(*
SPDX-FileCopyrightText: c 2026 Oleksandr Tiutyk <trofimich@gmail.com>
SPDX-License-Identifier: MIT
License: https://opensource.org/license/mit
*)

(*!
<summary>Groups fixed-capacity dictionary lookup, update, removal, clear and overflow cases.</summary>
<description>
Owns the child cases, their fixed registration array and the dictionaries borrowed by the common cases.
Each borrowed fixture is reserved for its case throughout the group lifetime. Use from one task at a stable address.
</description>
*)

{attribute 'no_assign'}
{attribute 'no_explicit_call' := 'do not call this function block directly'}
FUNCTION_BLOCK StaticDictionaryTestGroup EXTENDS TOF_Testing.TestGroup<5>
VAR_STAT
	{attribute 'hide'}
	_ClassName : STRING := __POUNAME();
END_VAR
VAR
	_SetAndGetDictionary : TOF_Collections.Dictionary<7>(keyValidator := 0, valueValidator := 0, keyEqualityComparer := 0);
	_RemoveDictionary : TOF_Collections.Dictionary<7>(keyValidator := 0, valueValidator := 0, keyEqualityComparer := 0);
	_ContainsDictionary : TOF_Collections.Dictionary<7>(keyValidator := 0, valueValidator := 0, keyEqualityComparer := 0);

	_SetAndGet : DictionarySetAndGetTest(name := "SetAndGet", parent := THIS^, dictionary := _SetAndGetDictionary);
	_Remove : DictionaryRemoveTest(name := "Remove", parent := THIS^, dictionary := _RemoveDictionary);
	_Contains : DictionaryContainsTest(name := "Contains", parent := THIS^, dictionary := _ContainsDictionary);
	_Clear : StaticDictionaryClearTest(name := "Clear", parent := THIS^);
	_Overflow : StaticDictionaryOverflowTest(name := "Overflow", parent := THIS^);

	_Children : ARRAY [0.._ChildCount - 1] OF TOF_Testing.ITestElement :=
	[
		_SetAndGet,
		_Remove,
		_Contains,
		_Clear,
		_Overflow
	];
END_VAR

//! <summary>Borrows the fixed child array. Callers must not modify it.</summary>
{attribute 'monitoring' := 'call'}
PROPERTY Children : REFERENCE TO ARRAY [0.._ChildCount - 1] OF TOF_Testing.ITestElement
GET
Children REF= _Children;
END_GET
END_PROPERTY

//! <summary>Borrows the concrete class name. Callers must not modify it.</summary>
{attribute 'monitoring' := 'call'}
PROPERTY ClassName : REFERENCE TO STRING
GET
ClassName REF= _ClassName;
END_GET
END_PROPERTY

//! <summary>Borrows the compiler-initialized namespace name. Callers must not modify it.</summary>
{attribute 'monitoring' := 'call'}
PROPERTY NamespaceName : REFERENCE TO STRING
GET
NamespaceName REF= CurrentNamespace.Name;
END_GET
END_PROPERTY

//! <summary>Reports the concrete instance size in bytes.</summary>
{attribute 'monitoring' := 'call'}
PROPERTY SelfSize : ULINT
GET
SelfSize := XSIZEOF(THIS^);
END_GET
END_PROPERTY

END_FUNCTION_BLOCK

(* stored: Version 1.1.0.1
   POU StaticDictionaryTestGroup: Id {3d8652fd-85fe-4723-aa37-3f2c000637c1}, SpecialFunc None
   Property Children: Id {355768cd-1f53-41e6-bd5c-894d10bb5e21}
   Get Get: Id {8be7babc-8716-4969-972c-11d36d526178}
   Property ClassName: Id {3d4da91e-07a1-4480-a20f-2011551f0e66}
   Get Get: Id {cfbc99c9-eeaa-44e7-8098-d5663cee2b28}
   Property NamespaceName: Id {1ac33c8f-139e-4285-b670-87d4eb3555d1}
   Get Get: Id {73f11067-5b0d-4079-97c3-0d64d5ca6bfb}
   Property SelfSize: Id {b37dcb3d-75aa-4da3-a363-dd24771e6430}
   Get Get: Id {a75d5ad3-c3ea-4f63-9109-232cd86abc06} *)
